Fanuc TP program (LS listing): Weld.LS

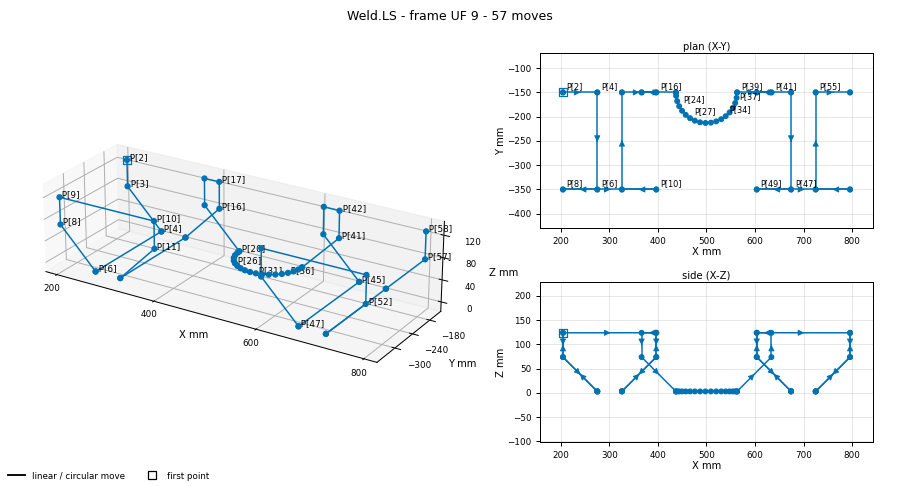
[picture p0: tool path of Weld.LS in frame UF 9, 57 of 58 moves have a stored position in this frame; points joined in program order, loops and branches not executed]
/PROG  Weld
/ATTR
OWNER		= MNEDITOR;
COMMENT		= "RoboDK sequence";
PROG_SIZE	= 0;
CREATE		= DATE 31-12-14  TIME 12:00:00;
MODIFIED	= DATE 31-12-14  TIME 12:00:00;
FILE_NAME	= Weld;
VERSION		= 0;
LINE_COUNT	= 83;
MEMORY_SIZE	= 0;
PROTECT		= READ_WRITE;
TCD:  STACK_SIZE	= 0,
      TASK_PRIORITY	= 50,
      TIME_SLICE	= 0,
      BUSY_LAMP_OFF	= 0,
      ABORT_REQUEST	= 0,
      PAUSE_REQUEST	= 0;
DEFAULT_GROUP	= 1,*,*,*,*,*,*;
CONTROL_CODE	= 00000000 00000000;
/MN
   1:  ! Program generated by VerticalBot Studio for Fanuc ARC Mate 12 ;
   2:  ! 0iB/10L on 25/10/2026 12:00:00 ;
   3:  ! Using nominal kinematics. ;
   4:  PR[9,1]=741.654 ;
   5:  PR[9,2]=-500.000 ;
   6:  PR[9,3]=-466.420 ;
   7:  PR[9,4]=0.000 ;
   8:  PR[9,5]=0.000 ;
   9:  PR[9,6]=90.000 ;
  10:  UFRAME[9]=PR[9] ;
  11:  UFRAME_NUM=9 ;
  12:  PR[9,1]=-2.000 ;
  13:  PR[9,2]=0.000 ;
  14:  PR[9,3]=402.000 ;
  15:  PR[9,4]=0.000 ;
  16:  PR[9,5]=45.000 ;
  17:  PR[9,6]=180.000 ;
  18:  UTOOL[9]=PR[9] ;
  19:  UTOOL_NUM=9 ;
  20:  ! show Daihen OTC weld gun ;
  21:J P[1] 20% CNT1 ;
  22:L P[2] 1000mm/sec CNT1 ;
  23:L P[3] 1000mm/sec CNT1 ;
  24:L P[4] 1000mm/sec FINE Arc Start[11] ;
  25:  Weave Sine[2.0Hz,8.0mm,0.075s,0.075] ;
  26:L P[5] 1000mm/sec CNT1 ;
  27:L P[6] 50mm/sec FINE Arc End[11] ;
  28:L P[7] 1000mm/sec CNT1 ;
  29:L P[8] 1000mm/sec CNT1 ;
  30:L P[9] 1000mm/sec CNT1 ;
  31:L P[10] 1000mm/sec CNT1 ;
  32:L P[11] 1000mm/sec CNT1 ;
  33:L P[12] 1000mm/sec FINE Arc Start[11] ;
  34:  Weave Sine[2.0Hz,8.0mm,0.075s,0.075] ;
  35:L P[13] 1000mm/sec CNT1 ;
  36:L P[14] 50mm/sec FINE Arc End[11] ;
  37:L P[15] 1000mm/sec CNT1 ;
  38:L P[16] 1000mm/sec CNT1 ;
  39:L P[17] 1000mm/sec CNT1 ;
  40:L P[18] 1000mm/sec CNT1 ;
  41:L P[19] 1000mm/sec CNT1 ;
  42:L P[20] 1000mm/sec FINE Arc Start[11] ;
  43:  Weave Sine[2.0Hz,8.0mm,0.075s,0.075] ;
  44:L P[21] 1000mm/sec CNT1 ;
  45:L P[22] 50mm/sec CNT1 ;
  46:L P[23] 50mm/sec CNT1 ;
  47:L P[24] 50mm/sec CNT1 ;
  48:L P[25] 50mm/sec CNT1 ;
  49:L P[26] 50mm/sec CNT1 ;
  50:L P[27] 50mm/sec CNT1 ;
  51:L P[28] 50mm/sec CNT1 ;
  52:L P[29] 50mm/sec CNT1 ;
  53:L P[30] 50mm/sec CNT1 ;
  54:L P[31] 50mm/sec CNT1 ;
  55:L P[32] 50mm/sec CNT1 ;
  56:L P[33] 50mm/sec CNT1 ;
  57:L P[34] 50mm/sec CNT1 ;
  58:L P[35] 50mm/sec CNT1 ;
  59:L P[36] 50mm/sec CNT1 ;
  60:L P[37] 50mm/sec CNT1 ;
  61:L P[38] 50mm/sec CNT1 ;
  62:L P[39] 50mm/sec FINE Arc End[11] ;
  63:L P[40] 1000mm/sec CNT1 ;
  64:L P[41] 1000mm/sec CNT1 ;
  65:L P[42] 1000mm/sec CNT1 ;
  66:L P[43] 1000mm/sec CNT1 ;
  67:L P[44] 1000mm/sec CNT1 ;
  68:L P[45] 1000mm/sec FINE Arc Start[11] ;
  69:  Weave Sine[2.0Hz,8.0mm,0.075s,0.075] ;
  70:L P[46] 1000mm/sec CNT1 ;
  71:L P[47] 50mm/sec FINE Arc End[11] ;
  72:L P[48] 1000mm/sec CNT1 ;
  73:L P[49] 1000mm/sec CNT1 ;
  74:L P[50] 1000mm/sec CNT1 ;
  75:L P[51] 1000mm/sec CNT1 ;
  76:L P[52] 1000mm/sec CNT1 ;
  77:L P[53] 1000mm/sec FINE Arc Start[11] ;
  78:  Weave Sine[2.0Hz,8.0mm,0.075s,0.075] ;
  79:L P[54] 1000mm/sec CNT1 ;
  80:L P[55] 50mm/sec FINE Arc End[11] ;
  81:L P[56] 1000mm/sec CNT1 ;
  82:L P[57] 1000mm/sec CNT1 ;
  83:L P[58] 1000mm/sec CNT1 ;
/POS
P[1]{
   GP1:
    UF : 9, UT : 9,
	J1=    -18.462 deg,	J2=    3.094 deg,	J3=    -45.099 deg,
	J4=    0.004 deg,	J5=    -44.900 deg,	J6=    -71.541 deg
};
P[2]{
   GP1:
    UF : 9, UT : 9,        CONFIG : 'F U T, 0, 0, 0',
	X =   204.293  mm,	Y =  -150.000  mm,	Z =   123.889  mm,
	W =   180.000 deg,	P =   -44.997 deg,	R =     0.000 deg
};
P[3]{
   GP1:
    UF : 9, UT : 9,        CONFIG : 'F U T, 0, 0, 0',
	X =   204.293  mm,	Y =  -150.000  mm,	Z =    73.889  mm,
	W =   180.000 deg,	P =   -44.997 deg,	R =     0.000 deg
};
P[4]{
   GP1:
    UF : 9, UT : 9,        CONFIG : 'F U T, 0, 0, 0',
	X =   275.000  mm,	Y =  -150.000  mm,	Z =     3.175  mm,
	W =   180.000 deg,	P =   -44.997 deg,	R =     0.000 deg
};
P[5]{
   GP1:
    UF : 9, UT : 9,        CONFIG : 'F U T, 0, 0, 0',
	X =   275.000  mm,	Y =  -150.000  mm,	Z =     3.175  mm,
	W =   180.000 deg,	P =   -44.997 deg,	R =     0.000 deg
};
P[6]{
   GP1:
    UF : 9, UT : 9,        CONFIG : 'F U T, 0, 0, 0',
	X =   275.000  mm,	Y =  -350.000  mm,	Z =     3.175  mm,
	W =  -180.000 deg,	P =   -44.997 deg,	R =     0.000 deg
};
P[7]{
   GP1:
    UF : 9, UT : 9,        CONFIG : 'F U T, 0, 0, 0',
	X =   275.000  mm,	Y =  -350.000  mm,	Z =     3.175  mm,
	W =  -180.000 deg,	P =   -44.997 deg,	R =     0.000 deg
};
P[8]{
   GP1:
    UF : 9, UT : 9,        CONFIG : 'F U T, 0, 0, 0',
	X =   204.293  mm,	Y =  -350.000  mm,	Z =    73.889  mm,
	W =  -180.000 deg,	P =   -44.997 deg,	R =     0.000 deg
};
P[9]{
   GP1:
    UF : 9, UT : 9,        CONFIG : 'F U T, 0, 0, 0',
	X =   204.293  mm,	Y =  -350.000  mm,	Z =   123.889  mm,
	W =  -180.000 deg,	P =   -44.997 deg,	R =     0.000 deg
};
P[10]{
   GP1:
    UF : 9, UT : 9,        CONFIG : 'F U T, 0, 0, 0',
	X =   396.511  mm,	Y =  -350.000  mm,	Z =   124.061  mm,
	W =  -161.118 deg,	P =   -41.641 deg,	R =   152.764 deg
};
P[11]{
   GP1:
    UF : 9, UT : 9,        CONFIG : 'F U T, 0, 0, 0',
	X =   396.511  mm,	Y =  -350.000  mm,	Z =    74.061  mm,
	W =   180.000 deg,	P =   -45.000 deg,	R =  -180.000 deg
};
P[12]{
   GP1:
    UF : 9, UT : 9,        CONFIG : 'F U T, 0, 0, 0',
	X =   325.800  mm,	Y =  -350.000  mm,	Z =     3.350  mm,
	W =   180.000 deg,	P =   -45.000 deg,	R =   180.000 deg
};
P[13]{
   GP1:
    UF : 9, UT : 9,        CONFIG : 'F U T, 0, 0, 0',
	X =   325.800  mm,	Y =  -350.000  mm,	Z =     3.350  mm,
	W =   180.000 deg,	P =   -45.000 deg,	R =  -180.000 deg
};
P[14]{
   GP1:
    UF : 9, UT : 9,        CONFIG : 'F U T, 0, 0, 0',
	X =   325.800  mm,	Y =  -150.000  mm,	Z =     3.350  mm,
	W =   180.000 deg,	P =   -45.000 deg,	R =   180.000 deg
};
P[15]{
   GP1:
    UF : 9, UT : 9,        CONFIG : 'F U T, 0, 0, 0',
	X =   325.800  mm,	Y =  -150.000  mm,	Z =     3.350  mm,
	W =   180.000 deg,	P =   -45.000 deg,	R =   180.000 deg
};
P[16]{
   GP1:
    UF : 9, UT : 9,        CONFIG : 'F U T, 0, 0, 0',
	X =   396.511  mm,	Y =  -150.000  mm,	Z =    74.061  mm,
	W =   180.000 deg,	P =   -45.000 deg,	R =  -180.000 deg
};
P[17]{
   GP1:
    UF : 9, UT : 9,        CONFIG : 'F U T, 0, 0, 0',
	X =   396.511  mm,	Y =  -150.000  mm,	Z =   124.061  mm,
	W =   180.000 deg,	P =   -45.000 deg,	R =  -180.000 deg
};
P[18]{
   GP1:
    UF : 9, UT : 9,        CONFIG : 'F U T, 0, 0, 1',
	X =   366.289  mm,	Y =  -150.000  mm,	Z =   123.886  mm,
	W =  -161.118 deg,	P =   -41.641 deg,	R =   -27.236 deg
};
P[19]{
   GP1:
    UF : 9, UT : 9,        CONFIG : 'F U T, 0, 0, 1',
	X =   366.289  mm,	Y =  -150.000  mm,	Z =    73.886  mm,
	W =  -180.000 deg,	P =   -45.000 deg,	R =     0.000 deg
};
P[20]{
   GP1:
    UF : 9, UT : 9,        CONFIG : 'F U T, 0, 0, 1',
	X =   437.000  mm,	Y =  -150.000  mm,	Z =     3.175  mm,
	W =   180.000 deg,	P =   -45.000 deg,	R =     0.000 deg
};
P[21]{
   GP1:
    UF : 9, UT : 9,        CONFIG : 'F U T, 0, 0, 1',
	X =   437.000  mm,	Y =  -150.000  mm,	Z =     3.175  mm,
	W =  -180.000 deg,	P =   -45.000 deg,	R =     0.000 deg
};
P[22]{
   GP1:
    UF : 9, UT : 9,        CONFIG : 'F U T, 0, 0, 1',
	X =   437.392  mm,	Y =  -157.018  mm,	Z =     3.175  mm,
	W =   180.000 deg,	P =   -45.000 deg,	R =     6.396 deg
};
P[23]{
   GP1:
    UF : 9, UT : 9,        CONFIG : 'F U T, 0, 0, 1',
	X =   439.628  mm,	Y =  -168.007  mm,	Z =     3.175  mm,
	W =  -180.000 deg,	P =   -45.000 deg,	R =    16.608 deg
};
P[24]{
   GP1:
    UF : 9, UT : 9,        CONFIG : 'F U T, 0, 0, 1',
	X =   443.777  mm,	Y =  -178.425  mm,	Z =     3.175  mm,
	W =   180.000 deg,	P =   -45.000 deg,	R =    26.820 deg
};
P[25]{
   GP1:
    UF : 9, UT : 9,        CONFIG : 'F U T, 0, 0, 1',
	X =   449.707  mm,	Y =  -187.942  mm,	Z =     3.175  mm,
	W =   180.000 deg,	P =   -45.000 deg,	R =    37.032 deg
};
P[26]{
   GP1:
    UF : 9, UT : 9,        CONFIG : 'F U T, 0, 0, 1',
	X =   457.231  mm,	Y =  -196.258  mm,	Z =     3.175  mm,
	W =  -180.000 deg,	P =   -45.000 deg,	R =    47.244 deg
};
P[27]{
   GP1:
    UF : 9, UT : 9,        CONFIG : 'F U T, 0, 0, 1',
	X =   466.109  mm,	Y =  -203.108  mm,	Z =     3.175  mm,
	W =   180.000 deg,	P =   -45.000 deg,	R =    57.456 deg
};
P[28]{
   GP1:
    UF : 9, UT : 9,        CONFIG : 'F U T, 0, 0, 1',
	X =   476.062  mm,	Y =  -208.275  mm,	Z =     3.175  mm,
	W =   180.000 deg,	P =   -45.000 deg,	R =    67.668 deg
};
P[29]{
   GP1:
    UF : 9, UT : 9,        CONFIG : 'F U T, 0, 0, 1',
	X =   486.772  mm,	Y =  -211.596  mm,	Z =     3.175  mm,
	W =   180.000 deg,	P =   -45.000 deg,	R =    77.880 deg
};
P[30]{
   GP1:
    UF : 9, UT : 9,        CONFIG : 'F U T, 0, 0, 1',
	X =   497.902  mm,	Y =  -212.965  mm,	Z =     3.175  mm,
	W =   180.000 deg,	P =   -45.000 deg,	R =    88.092 deg
};
P[31]{
   GP1:
    UF : 9, UT : 9,        CONFIG : 'F U T, 0, 0, 1',
	X =   509.099  mm,	Y =  -212.339  mm,	Z =     3.175  mm,
	W =   180.000 deg,	P =   -45.000 deg,	R =    98.304 deg
};
P[32]{
   GP1:
    UF : 9, UT : 9,        CONFIG : 'F U T, 0, 0, 1',
	X =   520.007  mm,	Y =  -209.739  mm,	Z =     3.175  mm,
	W =   180.000 deg,	P =   -45.000 deg,	R =   108.516 deg
};
P[33]{
   GP1:
    UF : 9, UT : 9,        CONFIG : 'F U T, 0, 0, 1',
	X =   530.281  mm,	Y =  -205.245  mm,	Z =     3.175  mm,
	W =   180.000 deg,	P =   -45.000 deg,	R =   118.728 deg
};
P[34]{
   GP1:
    UF : 9, UT : 9,        CONFIG : 'F U T, 0, 0, 1',
	X =   539.596  mm,	Y =  -199.002  mm,	Z =     3.175  mm,
	W =  -180.000 deg,	P =   -45.000 deg,	R =   128.940 deg
};
P[35]{
   GP1:
    UF : 9, UT : 9,        CONFIG : 'F U T, 0, 0, 1',
	X =   547.656  mm,	Y =  -191.205  mm,	Z =     3.175  mm,
	W =   180.000 deg,	P =   -45.000 deg,	R =   139.152 deg
};
P[36]{
   GP1:
    UF : 9, UT : 9,        CONFIG : 'F U T, 0, 0, 1',
	X =   554.207  mm,	Y =  -182.104  mm,	Z =     3.175  mm,
	W =   180.000 deg,	P =   -45.000 deg,	R =   149.364 deg
};
P[37]{
   GP1:
    UF : 9, UT : 9,        CONFIG : 'F U T, 0, 0, 1',
	X =   559.040  mm,	Y =  -171.985  mm,	Z =     3.175  mm,
	W =  -180.000 deg,	P =   -45.000 deg,	R =   159.576 deg
};
P[38]{
   GP1:
    UF : 9, UT : 9,        CONFIG : 'F U T, 0, 0, 1',
	X =   562.002  mm,	Y =  -161.169  mm,	Z =     3.175  mm,
	W =  -180.000 deg,	P =   -45.000 deg,	R =   169.788 deg
};
P[39]{
   GP1:
    UF : 9, UT : 9,        CONFIG : 'F U T, 0, 0, 1',
	X =   563.000  mm,	Y =  -150.000  mm,	Z =     3.175  mm,
	W =   180.000 deg,	P =   -45.000 deg,	R =  -180.000 deg
};
P[40]{
   GP1:
    UF : 9, UT : 9,        CONFIG : 'F U T, 0, 0, 1',
	X =   563.000  mm,	Y =  -150.000  mm,	Z =     3.175  mm,
	W =   180.000 deg,	P =   -45.000 deg,	R =  -180.000 deg
};
P[41]{
   GP1:
    UF : 9, UT : 9,        CONFIG : 'F U T, 0, 0, 1',
	X =   633.711  mm,	Y =  -150.000  mm,	Z =    73.886  mm,
	W =   180.000 deg,	P =   -45.000 deg,	R =  -180.000 deg
};
P[42]{
   GP1:
    UF : 9, UT : 9,        CONFIG : 'F U T, 0, 0, 1',
	X =   633.711  mm,	Y =  -150.000  mm,	Z =   123.886  mm,
	W =  -180.000 deg,	P =   -45.000 deg,	R =  -180.000 deg
};
P[43]{
   GP1:
    UF : 9, UT : 9,        CONFIG : 'F U T, 0, 0, 1',
	X =   603.489  mm,	Y =  -150.000  mm,	Z =   124.061  mm,
	W =   161.118 deg,	P =   -41.641 deg,	R =    27.236 deg
};
P[44]{
   GP1:
    UF : 9, UT : 9,        CONFIG : 'F U T, 0, 0, 1',
	X =   603.489  mm,	Y =  -150.000  mm,	Z =    74.061  mm,
	W =  -180.000 deg,	P =   -45.000 deg,	R =     0.000 deg
};
P[45]{
   GP1:
    UF : 9, UT : 9,        CONFIG : 'F U T, 0, 0, 1',
	X =   674.200  mm,	Y =  -150.000  mm,	Z =     3.350  mm,
	W =  -180.000 deg,	P =   -45.000 deg,	R =     0.000 deg
};
P[46]{
   GP1:
    UF : 9, UT : 9,        CONFIG : 'F U T, 0, 0, 1',
	X =   674.200  mm,	Y =  -150.000  mm,	Z =     3.350  mm,
	W =  -180.000 deg,	P =   -45.000 deg,	R =     0.000 deg
};
P[47]{
   GP1:
    UF : 9, UT : 9,        CONFIG : 'F U T, 0, 0, 1',
	X =   674.200  mm,	Y =  -350.000  mm,	Z =     3.350  mm,
	W =  -180.000 deg,	P =   -45.000 deg,	R =     0.000 deg
};
P[48]{
   GP1:
    UF : 9, UT : 9,        CONFIG : 'F U T, 0, 0, 1',
	X =   674.200  mm,	Y =  -350.000  mm,	Z =     3.350  mm,
	W =  -180.000 deg,	P =   -45.000 deg,	R =     0.000 deg
};
P[49]{
   GP1:
    UF : 9, UT : 9,        CONFIG : 'F U T, 0, 0, 1',
	X =   603.489  mm,	Y =  -350.000  mm,	Z =    74.061  mm,
	W =  -180.000 deg,	P =   -45.000 deg,	R =     0.000 deg
};
P[50]{
   GP1:
    UF : 9, UT : 9,        CONFIG : 'F U T, 0, 0, 1',
	X =   603.489  mm,	Y =  -350.000  mm,	Z =   124.061  mm,
	W =  -180.000 deg,	P =   -45.000 deg,	R =     0.000 deg
};
P[51]{
   GP1:
    UF : 9, UT : 9,        CONFIG : 'F U T, 0, 0, 1',
	X =   795.711  mm,	Y =  -350.000  mm,	Z =   123.886  mm,
	W =  -161.118 deg,	P =   -41.641 deg,	R =   152.764 deg
};
P[52]{
   GP1:
    UF : 9, UT : 9,        CONFIG : 'F U T, 0, 0, 1',
	X =   795.711  mm,	Y =  -350.000  mm,	Z =    73.886  mm,
	W =   180.000 deg,	P =   -45.000 deg,	R =  -180.000 deg
};
P[53]{
   GP1:
    UF : 9, UT : 9,        CONFIG : 'F U T, 0, 0, 1',
	X =   725.000  mm,	Y =  -350.000  mm,	Z =     3.175  mm,
	W =   180.000 deg,	P =   -45.000 deg,	R =   180.000 deg
};
P[54]{
   GP1:
    UF : 9, UT : 9,        CONFIG : 'F U T, 0, 0, 1',
	X =   725.000  mm,	Y =  -350.000  mm,	Z =     3.175  mm,
	W =   180.000 deg,	P =   -45.000 deg,	R =   180.000 deg
};
P[55]{
   GP1:
    UF : 9, UT : 9,        CONFIG : 'F U T, 0, 0, 1',
	X =   725.000  mm,	Y =  -150.000  mm,	Z =     3.175  mm,
	W =   180.000 deg,	P =   -45.000 deg,	R =  -180.000 deg
};
P[56]{
   GP1:
    UF : 9, UT : 9,        CONFIG : 'F U T, 0, 0, 1',
	X =   725.000  mm,	Y =  -150.000  mm,	Z =     3.175  mm,
	W =   180.000 deg,	P =   -45.000 deg,	R =  -180.000 deg
};
P[57]{
   GP1:
    UF : 9, UT : 9,        CONFIG : 'F U T, 0, 0, 1',
	X =   795.711  mm,	Y =  -150.000  mm,	Z =    73.886  mm,
	W =   180.000 deg,	P =   -45.000 deg,	R =   180.000 deg
};
P[58]{
   GP1:
    UF : 9, UT : 9,        CONFIG : 'F U T, 0, 0, 1',
	X =   795.711  mm,	Y =  -150.000  mm,	Z =   123.886  mm,
	W =  -180.000 deg,	P =   -45.000 deg,	R =   180.000 deg
};
/END
